(* IEC 61131-3 sources: PLC_ST_Auto/tests/llm_eval_golden, 14 files *)

(* ---- TC-01.st ---- *)
PROGRAM MotorStartStop
VAR_INPUT
    start : BOOL; (* Start pushbutton, normally-open contact, TRUE = pressed *)
    stop  : BOOL; (* Stop pushbutton, TRUE = pressed *)
                  (* Assumption: stop is wired as a normally-open signal.
                     If a normally-closed stop button is used (the usual
                     fail-safe wiring), invert this signal before it is
                     connected to this program. *)
END_VAR
VAR_OUTPUT
    motor : BOOL; (* Contactor output *)
END_VAR

(* Seal-in (latching) circuit: the motor output is its own holding contact.
   The stop condition is ANDed last, so stop always has priority:
   if start and stop are pressed together, motor stays OFF. *)
motor := (start OR motor) AND NOT stop;

END_PROGRAM

(* ---- TC-02.st ---- *)
PROGRAM StarDeltaStarter
VAR_INPUT
    start : BOOL;   (* Start pushbutton, momentary NO *)
    stop  : BOOL;   (* Stop input, TRUE = stop request; stop has priority *)
END_VAR
VAR_OUTPUT
    km_main  : BOOL; (* Main contactor *)
    km_star  : BOOL; (* Star contactor *)
    km_delta : BOOL; (* Delta contactor *)
END_VAR
VAR
    running   : BOOL;  (* Latched run command *)
    tmr_star  : TON;   (* Star running time: 5000 ms *)
    tmr_dead  : TON;   (* Star-to-delta dead time *)
END_VAR

(* Assumptions:
   - start is a momentary pushbutton, so the run command is latched internally.
   - stop is TRUE when a stop is requested. If a normally closed stop button is used,
     invert it at the input mapping.
   - A 100 ms dead time between km_star dropping out and km_delta pulling in
     is added as extra protection against short circuit (contactor arc/off delay).
   - No overload input was specified, so none is implemented. *)

(* Run latch, stop priority *)
running := (start OR running) AND NOT stop;

(* Star time of 5 s, started when running *)
tmr_star(IN := running, PT := T#5000ms);

(* Dead time starts when the star time has elapsed *)
tmr_dead(IN := running AND tmr_star.Q, PT := T#100ms);

(* Main contactor *)
km_main := running;

(* Star contactor: only during the star phase, interlocked with delta *)
km_star := running AND NOT tmr_star.Q AND NOT km_delta;

(* Delta contactor: after dead time, interlocked with star *)
km_delta := running AND tmr_dead.Q AND NOT km_star;

END_PROGRAM

(* ---- TC-03.st ---- *)
PROGRAM PackageCounter
VAR_INPUT
    sensor    : BOOL;   (* Photoelectric sensor: TRUE while a workpiece is detected *)
    reset_btn : BOOL;   (* Reset pushbutton: TRUE while pressed *)
END_VAR
VAR_OUTPUT
    package_ready : BOOL;  (* TRUE when the count reaches the package quantity *)
    count_value   : INT;   (* Current accumulated count, for display/monitoring *)
END_VAR
VAR
    cnt_ctu : CTU;         (* Standard IEC up-counter *)
    PACK_QTY : INT := 10;  (* Preset package quantity *)
END_VAR

(* Assumptions:
   - The CTU counts rising edges on its CU input internally (it contains an R_TRIG),
     so each workpiece passing is counted once per rising edge of sensor.
   - While reset_btn is TRUE, R is dominant: the counter is cleared to 0
     and package_ready (Q) is FALSE.
   - After reaching PV the CTU keeps counting further pulses and Q stays TRUE
     until reset; package_ready therefore stays latched until reset_btn is pressed. *)

cnt_ctu(CU := sensor,
        R  := reset_btn,
        PV := PACK_QTY);

package_ready := cnt_ctu.Q;
count_value   := cnt_ctu.CV;

END_PROGRAM

(* ---- TC-04.st ---- *)
PROGRAM TrafficLight
VAR_INPUT
    emergency : BOOL;   (* TRUE = force all-red mode immediately *)
END_VAR
VAR_OUTPUT
    green  : BOOL;
    yellow : BOOL;
    red    : BOOL;
END_VAR
VAR
    State      : INT := 0;      (* 0=green, 1=yellow, 2=red *)
    tGreen     : TON;
    tYellow    : TON;
    tRed       : TON;
END_VAR

(* Assumptions:
   - While emergency is TRUE: only red is ON, all timers are reset.
   - When emergency is released, the cycle restarts from State 0 (green)
     with a fresh 5 s timer.
   - Each state's timer runs only while that state is active. *)

IF emergency THEN
    State := 0;   (* restart cycle from green after emergency is cleared *)
    tGreen(IN := FALSE, PT := T#5s);
    tYellow(IN := FALSE, PT := T#2s);
    tRed(IN := FALSE, PT := T#5s);
    green  := FALSE;
    yellow := FALSE;
    red    := TRUE;
ELSE
    tGreen(IN := (State = 0), PT := T#5s);
    tYellow(IN := (State = 1), PT := T#2s);
    tRed(IN := (State = 2), PT := T#5s);

    CASE State OF
        0:  (* Green *)
            green  := TRUE;
            yellow := FALSE;
            red    := FALSE;
            IF tGreen.Q THEN
                State := 1;
            END_IF;

        1:  (* Yellow *)
            green  := FALSE;
            yellow := TRUE;
            red    := FALSE;
            IF tYellow.Q THEN
                State := 2;
            END_IF;

        2:  (* Red *)
            green  := FALSE;
            yellow := FALSE;
            red    := TRUE;
            IF tRed.Q THEN
                State := 0;
            END_IF;

    ELSE
        (* Invalid state: recover to green *)
        State := 0;
        green  := FALSE;
        yellow := FALSE;
        red    := TRUE;
    END_CASE;
END_IF;

END_PROGRAM

(* ---- TC-05.st ---- *)
PROGRAM water_tank_control
VAR_INPUT
  emergency_stop : BOOL := false; (* 現場急停開關 *)
  high_level_sw : BOOL := false; (* 水槽高水位浮球 *)
  low_level_sw : BOOL := false; (* 水槽低水位浮球 *)
END_VAR
VAR_OUTPUT
  inlet_valve : BOOL := false; (* 進水電磁閥 *)
  drain_pump : BOOL := false; (* 排水泵浦 *)
  alarm_lamp : BOOL := false; (* 水位警報燈 *)
END_VAR
VAR
  fill_time : TIME := T#0s; (* 進水累計時間 *)
  fill_timer : TON;
END_VAR

(* Assumptions:
   - emergency_stop = TRUE means emergency active (TRUE = stop requested).
   - low_level_sw = TRUE means water is at or below the low level.
   - high_level_sw = TRUE means water is at or above the high level.
   - Inlet valve latches on at low level and stays on until high level
     (the requirement does not specify the hold behaviour).
   - Drain pump starts at high level and stops when low level is reached
     (stop condition is not specified in the requirement).
   - fill_time shows the elapsed time of the current filling run and
     resets to 0 when the inlet valve closes (TON elapsed time, max 1 h). *)

IF emergency_stop THEN
  (* Emergency: everything off, alarm lamp on *)
  inlet_valve := FALSE;
  drain_pump  := FALSE;
  alarm_lamp  := TRUE;
ELSE
  alarm_lamp := FALSE;

  IF high_level_sw THEN
    (* High level: close inlet, start drain pump *)
    inlet_valve := FALSE;
    drain_pump  := TRUE;
  ELSIF low_level_sw THEN
    (* Low level and not high: open inlet, stop pump *)
    inlet_valve := TRUE;
    drain_pump  := FALSE;
  ELSE
    (* Between levels: keep previous state (hysteresis);
       inlet and pump are never on at the same time *)
    IF inlet_valve AND drain_pump THEN
      inlet_valve := FALSE;
    END_IF;
  END_IF;
END_IF;

(* Fill time measurement *)
fill_timer(IN := inlet_valve, PT := T#1h);
fill_time := fill_timer.ET;

END_PROGRAM

(* ---- TC-06.st ---- *)
PROGRAM AnalogMovingAvg5
VAR_INPUT
    raw_in : REAL;                      (* raw analog value *)
END_VAR
VAR_OUTPUT
    filter_out : REAL;                  (* filtered output *)
END_VAR
VAR
    buf : ARRAY[0..4] OF REAL := [0.0, 0.0, 0.0, 0.0, 0.0];  (* last 5 samples *)
    idx : INT := 0;                     (* write index 0..4 *)
    i   : INT;
    sum : REAL;
END_VAR

(* Assumption: the buffer starts at 0.0, so during the first 4 scans
   the average includes these initial zeros, as the standard's algorithm
   (sum of 5 points / 5.0) specifies. *)

(* Safety guard: keep the index within the valid range *)
IF (idx < 0) OR (idx > 4) THEN
    idx := 0;
END_IF;

(* Write the new sample into the buffer *)
buf[idx] := raw_in;

(* Sum the 5 points *)
sum := 0.0;
FOR i := 0 TO 4 DO
    sum := sum + buf[i];
END_FOR;

(* Moving average *)
filter_out := sum / 5.0;

(* Advance the circular index *)
idx := (idx + 1) MOD 5;

END_PROGRAM

(* ---- TC-07.st ---- *)
PROGRAM TempControl
VAR_INPUT
    temp_pv : REAL;   (* Process value (analog input, engineering units) *)
    temp_sp : REAL;   (* Setpoint *)
END_VAR
VAR_OUTPUT
    heater : BOOL;    (* Heater output *)
    cooler : BOOL;    (* Cooler output *)
END_VAR
VAR
    hyst : REAL := 2.0;   (* Hysteresis band +/- 2.0 around setpoint *)
END_VAR

(* Assumptions:
   - Inside the dead band (sp-2.0 <= pv <= sp+2.0) the outputs hold their
     previous state (latching on/off hysteresis behaviour), since the
     requirement does not specify otherwise.
   - Heater is switched off when the cooler is started (pv > sp+2.0).
   - Cooler is switched off when the heater is started (pv < sp-2.0).
     This guarantees heater and cooler are never on simultaneously.
   - Cooler stays on until the temperature falls below sp-2.0 (heating
     demand); heater stays on until pv exceeds sp+2.0. Adjust here if
     a different switch-off point (e.g. at setpoint) is desired. *)

IF temp_pv < (temp_sp - hyst) THEN
    heater := TRUE;
    cooler := FALSE;
ELSIF temp_pv > (temp_sp + hyst) THEN
    heater := FALSE;
    cooler := TRUE;
END_IF;

END_PROGRAM

(* ---- TC-08.st ---- *)
PROGRAM Conveyor_Control
VAR_INPUT
    start        : BOOL;   (* 啟動按鈕 (常開, 按下=TRUE) *)
    stop         : BOOL;   (* 停止按鈕 (假設為常開, 按下=TRUE; 若為常閉接線請於輸入映射時反相) *)
    item_trigger : BOOL;   (* 光電開關, 物件通過時為 TRUE *)
    count_reset  : BOOL;   (* 產量歸零按鈕 (額外提供, 非必要) *)
END_VAR
VAR_OUTPUT
    conveyor     : BOOL;   (* 輸送帶馬達運轉輸出 *)
    item_count   : DINT;   (* 累計產量 *)
END_VAR
VAR
    run_latch    : BOOL;   (* 運轉自保持 *)
    trig_item    : R_TRIG; (* 光電開關上升緣偵測, 避免同一物件重複計數 *)
END_VAR

(* 假設: 停止優先於啟動; 僅在輸送帶運轉時才累計產量 *)
run_latch := (start OR run_latch) AND NOT stop;
conveyor  := run_latch;

(* 光電開關上升緣偵測 *)
trig_item(CLK := item_trigger);

IF count_reset THEN
    item_count := 0;
ELSIF trig_item.Q AND run_latch THEN
    IF item_count < 2147483647 THEN   (* 防止 DINT 溢位 *)
        item_count := item_count + 1;
    END_IF;
END_IF;

END_PROGRAM

(* ---- TC-09.st ---- *)
PROGRAM DualMotorSequence
VAR_INPUT
    start : BOOL;
    stop  : BOOL;
END_VAR
VAR_OUTPUT
    motor1 : BOOL;
    motor2 : BOOL;
END_VAR
VAR
    delay2 : TON;
END_VAR
(* Assumption: start is momentary; stop has priority *)
motor1 := (start OR motor1) AND NOT stop;
delay2(IN := motor1, PT := T#3s);
motor2 := motor1 AND delay2.Q;
END_PROGRAM

(* ---- TC-10.st ---- *)
PROGRAM PumpStartStop
VAR_INPUT
    start : BOOL;   (* Start pushbutton, normally open: TRUE = pressed *)
    stop  : BOOL;   (* Stop pushbutton: TRUE = pressed (assumption: NO contact, no fail-safe wiring) *)
END_VAR
VAR_OUTPUT
    pump      : BOOL;  (* Pump contactor command *)
    run_hours : INT;   (* Accumulated full running hours; held at 32767 max *)
END_VAR
VAR
    pump_latch : BOOL := FALSE;
    hour_timer : TON;
END_VAR

(* Classic seal-in circuit; stop has priority over start *)
pump_latch := (start OR pump_latch) AND NOT stop;
pump := pump_latch;

(* Run-hour counter: 1 h timer runs only while pump is on.
   Assumption: partial hours are lost when the pump stops (timer resets);
   run_hours is not retentive across power cycles unless the vendor makes it so. *)
hour_timer(IN := pump_latch AND NOT hour_timer.Q, PT := T#1h);

IF hour_timer.Q THEN
    IF run_hours < 32767 THEN
        run_hours := run_hours + 1;
    END_IF;
END_IF;

END_PROGRAM

(* ---- TC-11.st ---- *)
PROGRAM FireAlarmSystem
VAR_INPUT
    fire_sensor : BOOL;   (* TRUE = fire detected *)
    ack_btn     : BOOL;   (* acknowledge push button *)
END_VAR
VAR_OUTPUT
    alarm : BOOL;         (* alarm output, latched *)
    siren : BOOL;         (* buzzer output, latched *)
END_VAR
VAR
    tmr_siren : TON;
    ack_edge  : R_TRIG;
END_VAR

(* Assumptions:
   - alarm and siren are latched: they stay TRUE even if the fire signal
     disappears, until the fire is cleared AND ack_btn is pressed.
   - Acknowledge is evaluated on the rising edge of ack_btn, and only
     when fire_sensor is FALSE at that moment.
   - If fire_sensor is active again, the alarm is set again immediately
     (fire has priority over reset).
   - The 400 ms timer runs only while fire_sensor is continuously TRUE;
     siren is latched once the timer elapses. *)

(* Siren delay timer: fire continuously present for 400 ms *)
tmr_siren(IN := fire_sensor, PT := T#400ms);

(* Acknowledge button edge detection *)
ack_edge(CLK := ack_btn);

(* Set: alarm immediately on fire *)
IF fire_sensor THEN
    alarm := TRUE;
END_IF;

(* Set: siren after fire lasted more than 400 ms *)
IF tmr_siren.Q THEN
    siren := TRUE;
END_IF;

(* Reset: fire cleared and acknowledge pressed (fire has priority) *)
IF ack_edge.Q AND NOT fire_sensor THEN
    alarm := FALSE;
    siren := FALSE;
END_IF;

END_PROGRAM

(* ---- TC-12.st ---- *)
PROGRAM HighSpeedProductionCounter
VAR_INPUT
    pulse : BOOL;   (* Sensor pulse input *)
    clear : BOOL;   (* Reset button: clears total_count to 0 *)
END_VAR
VAR_OUTPUT
    total_count : INT := 0;        (* Total production count, saturates at 32767 *)
    at_limit    : BOOL := FALSE;   (* TRUE when counter has reached the upper limit *)
END_VAR
VAR
    pulse_trig : R_TRIG;   (* Rising edge detector for pulse *)
END_VAR

(* Assumption: clear has priority over counting when both occur in the same scan. *)
(* Assumption: the rising edge detection is evaluated every scan; the pulse must be
   slower than the PLC scan time to be captured (a true high-speed input would require
   a hardware counter, which is outside standard IEC ST). *)

pulse_trig(CLK := pulse);

IF clear THEN
    total_count := 0;
ELSIF pulse_trig.Q THEN
    IF total_count < 32767 THEN
        total_count := total_count + 1;
    END_IF;
END_IF;

at_limit := (total_count >= 32767);

END_PROGRAM

(* ---- TC-13.st ---- *)
PROGRAM FAN_CONTROL
VAR_INPUT
    run_cmd  : BOOL; (* Start pushbutton, normally open *)
    stop_cmd : BOOL; (* Stop command; assumption: TRUE = stop requested *)
END_VAR
VAR_OUTPUT
    fan_out  : BOOL; (* Fan contactor output *)
END_VAR
VAR
    fan_latch : BOOL; (* Internal seal-in memory *)
END_VAR

(* Assumptions:
   - Stop has priority over run (safety): if both buttons are pressed
     at the same time, the fan is stopped / stays off.
   - stop_cmd is treated as active-high (TRUE = stop pressed).
     For a wiring-fault-safe design, a normally-closed stop button
     would normally be used and inverted here.
   - The fan does not automatically restart after both buttons are
     released, because the stop command resets the latch; a new
     rising run_cmd with stop_cmd = FALSE is required.
   - Latch is not retained, so fan is off after power-up. *)

(* Stop-dominant seal-in logic *)
fan_latch := (run_cmd OR fan_latch) AND NOT stop_cmd;

fan_out := fan_latch;

END_PROGRAM

(* ---- TC-14.st ---- *)
PROGRAM CoolingTower
VAR_INPUT
    start : BOOL;
    stop  : BOOL;
END_VAR
VAR_OUTPUT
    pump : BOOL;
END_VAR
pump := (start OR pump) AND NOT stop;
END_PROGRAM
